// The stop is held until the stop transaction has settled (3A.2).
METHOD PRIVATE Stop_Is_Held_Until_The_Transaction_Settles
VAR_INST
	rig			: FB_IagRig;
	nStep		: INT;
	nCycles		: UINT;
	nEdges		: UINT;
	bSeen		: BOOL;
	sTest		: STRING(80);
END_VAR
TEST('Stop_Is_Held_Until_The_Transaction_Settles');
sTest := 'Stop_Is_Held_Until_The_Transaction_Settles: ';
IF nStep >= 90 THEN
	RETURN;
END_IF
rig.Scan();
nCycles := nCycles + 1;
CASE nStep OF
0:	// wait for the clock, then power on
	IF rig.ClockValid THEN
		rig.fbTel.Init();
		nStep := 10;
		nCycles := 0;
	ELSIF nCycles > 2000 THEN
		AssertTrue(Condition := FALSE, Message := 'the astronomical clock never became valid');
		F_Note(bFailed := TRUE, sText := CONCAT(sTest, 'the astronomical clock never became valid'));
		nStep := 99;
		TEST_FINISHED();
	END_IF
10:	// wait until the startup has finished (READY_STATE 1.0)
	IF rig.Online THEN
		rig.fbTel.Slew(fAzimuth := 180.0, fAltitude := 45.0);
		nStep := 20;
		nCycles := 0;
	ELSIF nCycles > 1500 THEN
		AssertTrue(Condition := FALSE, Message := 'the mock telescope did not reach READY_STATE 1.0');
		F_Note(bFailed := TRUE, sText := CONCAT(sTest, 'the mock telescope did not reach READY_STATE 1.0'));
		nStep := 99;
		TEST_FINISHED();
	END_IF
20:	// an axis is moving
	IF rig.fbHa.MoveAxis OR rig.fbDec.MoveAxis THEN
		nCycles := 0;
		nStep := 30;
	ELSIF nCycles > 300 THEN
		AssertTrue(Condition := FALSE, Message := 'the slew did not start an axis move');
		F_Note(bFailed := TRUE, sText := CONCAT(sTest, 'the slew did not start an axis move'));
		nStep := 99;
		TEST_FINISHED();
	END_IF
30:
	IF nCycles >= 5 THEN
		rig.fbTel.Stop();
		nStep := 40;
		nCycles := 0;
	END_IF
40:	// the stop is held while the axis is stopping, and released only when the transaction has settled
	IF nCycles = 2 THEN
		AssertTrue(Condition := rig.fbTel.bStopActive, Message := 'the stop is still held two scans after the command');
		F_Note(bFailed := NOT (rig.fbTel.bStopActive), sText := CONCAT(sTest, 'the stop is still held two scans after the command'));
	END_IF
	IF NOT rig.fbTel.bStopActive THEN
		AssertTrue(Condition := rig.fbTel.bSettled, Message := 'released only when settled');
		F_Note(bFailed := NOT (rig.fbTel.bSettled), sText := CONCAT(sTest, 'released only when settled'));
		nStep := 99;
		TEST_FINISHED();
	ELSIF nCycles > 400 THEN
		AssertTrue(Condition := FALSE, Message := 'the stop did not settle');
		F_Note(bFailed := TRUE, sText := CONCAT(sTest, 'the stop did not settle'));
		nStep := 99;
		TEST_FINISHED();
	END_IF
END_CASE
END_METHOD

// A goto and a home that are both pending when the stop comes are both cleared (3A.3).
METHOD PRIVATE Stop_Clears_Every_Pending_Move
VAR_INST
	rig			: FB_IagRig;
	nStep		: INT;
	nCycles		: UINT;
	nEdges		: UINT;
	bSeen		: BOOL;
	sTest		: STRING(80);
END_VAR
TEST('Stop_Clears_Every_Pending_Move');
sTest := 'Stop_Clears_Every_Pending_Move: ';
IF nStep >= 90 THEN
	RETURN;
END_IF
rig.Scan();
nCycles := nCycles + 1;
CASE nStep OF
0:	// wait for the clock, then power on
	IF rig.ClockValid THEN
		rig.fbTel.Init();
		nStep := 10;
		nCycles := 0;
	ELSIF nCycles > 2000 THEN
		AssertTrue(Condition := FALSE, Message := 'the astronomical clock never became valid');
		F_Note(bFailed := TRUE, sText := CONCAT(sTest, 'the astronomical clock never became valid'));
		nStep := 99;
		TEST_FINISHED();
	END_IF
10:	// wait until the startup has finished (READY_STATE 1.0)
	IF rig.Online THEN
		rig.fbTel.Track(fRightAscension := 100.0, fDeclination := 30.0);
		rig.fbTel.Home();
		rig.fbTel.Stop();
		nStep := 20;
		nCycles := 0;
	ELSIF nCycles > 1500 THEN
		AssertTrue(Condition := FALSE, Message := 'the mock telescope did not reach READY_STATE 1.0');
		F_Note(bFailed := TRUE, sText := CONCAT(sTest, 'the mock telescope did not reach READY_STATE 1.0'));
		nStep := 99;
		TEST_FINISHED();
	END_IF
20:	// one scan after the three commands
		AssertTrue(Condition := NOT rig.fbTel.bGotoActive, Message := 'the goto is gone');
		F_Note(bFailed := NOT (NOT rig.fbTel.bGotoActive), sText := CONCAT(sTest, 'the goto is gone'));
		AssertTrue(Condition := NOT rig.fbTel.bGoHomeActive, Message := 'the home is gone');
		F_Note(bFailed := NOT (NOT rig.fbTel.bGoHomeActive), sText := CONCAT(sTest, 'the home is gone'));
		nStep := 99;
		TEST_FINISHED();
END_CASE
END_METHOD

// A repeated stop does not send a second stop to an axis that is already stopping (3A.4).
METHOD PRIVATE Repeated_Stop_Restarts_Only_Moving_Axes
VAR_INST
	rig			: FB_IagRig;
	nStep		: INT;
	nCycles		: UINT;
	nEdges		: UINT;
	bSeen		: BOOL;
	sTest		: STRING(80);
END_VAR
TEST('Repeated_Stop_Restarts_Only_Moving_Axes');
sTest := 'Repeated_Stop_Restarts_Only_Moving_Axes: ';
IF nStep >= 90 THEN
	RETURN;
END_IF
rig.Scan();
nCycles := nCycles + 1;
CASE nStep OF
0:	// wait for the clock, then power on
	IF rig.ClockValid THEN
		rig.fbTel.Init();
		nStep := 10;
		nCycles := 0;
	ELSIF nCycles > 2000 THEN
		AssertTrue(Condition := FALSE, Message := 'the astronomical clock never became valid');
		F_Note(bFailed := TRUE, sText := CONCAT(sTest, 'the astronomical clock never became valid'));
		nStep := 99;
		TEST_FINISHED();
	END_IF
10:	// wait until the startup has finished (READY_STATE 1.0)
	IF rig.Online THEN
		rig.fbTel.Slew(fAzimuth := 180.0, fAltitude := 45.0);
		nStep := 20;
		nCycles := 0;
	ELSIF nCycles > 1500 THEN
		AssertTrue(Condition := FALSE, Message := 'the mock telescope did not reach READY_STATE 1.0');
		F_Note(bFailed := TRUE, sText := CONCAT(sTest, 'the mock telescope did not reach READY_STATE 1.0'));
		nStep := 99;
		TEST_FINISHED();
	END_IF
20:	// an axis is moving
	IF rig.fbHa.MoveAxis OR rig.fbDec.MoveAxis THEN
		nCycles := 0;
		nStep := 30;
	ELSIF nCycles > 300 THEN
		AssertTrue(Condition := FALSE, Message := 'the slew did not start an axis move');
		F_Note(bFailed := TRUE, sText := CONCAT(sTest, 'the slew did not start an axis move'));
		nStep := 99;
		TEST_FINISHED();
	END_IF
30:
	IF nCycles >= 5 THEN
		rig.fbTel.Stop();
		nStep := 35;
		nCycles := 0;
	END_IF
35:	// a second stop while the axis is already stopping (the stop reaches the axis in the third scan, the axis then reports Stopping)
	IF nCycles >= 3 THEN
		rig.fbTel.Stop();
		nStep := 40;
		nCycles := 0;
	END_IF
40:
	IF NOT rig.fbTel.bStopActive AND rig.fbTel.bStopped AND nCycles > 5 THEN
		AssertTrue(Condition := rig.fbHa.nStopEdges + rig.fbDec.nStopEdges = 1, Message := 'no second stop for an axis that was stopping');
		F_Note(bFailed := NOT (rig.fbHa.nStopEdges + rig.fbDec.nStopEdges = 1), sText := CONCAT(sTest, 'no second stop for an axis that was stopping'));
		nStep := 99;
		TEST_FINISHED();
	ELSIF nCycles > 400 THEN
		AssertTrue(Condition := FALSE, Message := 'the stop did not settle');
		F_Note(bFailed := TRUE, sText := CONCAT(sTest, 'the stop did not settle'));
		nStep := 99;
		TEST_FINISHED();
	END_IF
END_CASE
END_METHOD

// A park over a goto that is not dispatched yet runs a short abort stop, then the park (3A.5).
METHOD PRIVATE Park_Over_A_Waiting_Goto_Runs_A_Short_Abort_Stop
VAR_INST
	rig			: FB_IagRig;
	nStep		: INT;
	nCycles		: UINT;
	nEdges		: UINT;
	bSeen		: BOOL;
	sTest		: STRING(80);
END_VAR
TEST('Park_Over_A_Waiting_Goto_Runs_A_Short_Abort_Stop');
sTest := 'Park_Over_A_Waiting_Goto_Runs_A_Short_Abort_Stop: ';
IF nStep >= 90 THEN
	RETURN;
END_IF
rig.Scan();
nCycles := nCycles + 1;
CASE nStep OF
0:	// wait for the clock, then power on
	IF rig.ClockValid THEN
		rig.fbTel.Init();
		nStep := 10;
		nCycles := 0;
	ELSIF nCycles > 2000 THEN
		AssertTrue(Condition := FALSE, Message := 'the astronomical clock never became valid');
		F_Note(bFailed := TRUE, sText := CONCAT(sTest, 'the astronomical clock never became valid'));
		nStep := 99;
		TEST_FINISHED();
	END_IF
10:	// wait until the startup has finished (READY_STATE 1.0)
	IF rig.Online THEN
		rig.SetHorizon(-90.0);
		rig.SetSafeAltitude(-90.0);
		rig.fbTel.Track(fRightAscension := 100.0, fDeclination := 30.0);
		rig.fbTel.Park();
		nStep := 20;
		nCycles := 0;
	ELSIF nCycles > 1500 THEN
		AssertTrue(Condition := FALSE, Message := 'the mock telescope did not reach READY_STATE 1.0');
		F_Note(bFailed := TRUE, sText := CONCAT(sTest, 'the mock telescope did not reach READY_STATE 1.0'));
		nStep := 99;
		TEST_FINISHED();
	END_IF
20:	// the park preempted a goto that was not dispatched: the abort stop runs, then the park
	IF rig.fbTel.bMoveAbortPending THEN
		bSeen := TRUE;
	END_IF
	IF rig.fbTel.bIsParked THEN
		AssertTrue(Condition := bSeen, Message := 'the preemption ran the abort stop');
		F_Note(bFailed := NOT (bSeen), sText := CONCAT(sTest, 'the preemption ran the abort stop'));
		AssertTrue(Condition := NOT rig.fbTel.bGotoActive, Message := 'the goto is gone');
		F_Note(bFailed := NOT (NOT rig.fbTel.bGotoActive), sText := CONCAT(sTest, 'the goto is gone'));
		nStep := 99;
		TEST_FINISHED();
	ELSIF nCycles > 3000 THEN
		AssertTrue(Condition := FALSE, Message := 'the park did not finish');
		F_Note(bFailed := TRUE, sText := CONCAT(sTest, 'the park did not finish'));
		nStep := 99;
		TEST_FINISHED();
	END_IF
END_CASE
END_METHOD

END_FUNCTION_BLOCK

// ---- POUs/IagParkPowerReset_Tests.TcPOU
// Park, power-on and reset precedence of FB_TelescopeControl (IAG50cm), command model step 3B (BROTLib
// specs/plans/2026-11-09-iag50cm-command-model-unification.md). One rig per test, one Scan() per PLC cycle.
FUNCTION_BLOCK IagParkPowerReset_Tests EXTENDS TcUnit.FB_TestSuite
VAR
END_VAR

Park_During_Stop_Runs_After_Settle();
Stop_Drops_A_Park_Queued_Behind_A_Stop();
Init_During_Stop_Is_Refused();
Init_During_Park_Is_Refused();
Park_Right_After_Init_Aborts_The_PowerOn();
Init_Drops_A_Stale_Home();
Reset_At_Rest_Drops_A_Pending_Move();
Reset_During_Park_Keeps_The_Park();
Reset_Recovers_A_Stuck_Stop();

// A park sent during a stop runs when the stop has settled (D13).
METHOD PRIVATE Park_During_Stop_Runs_After_Settle
VAR_INST
	rig			: FB_IagRig;
	nStep		: INT;
	nCycles		: UINT;
	bSeen		: BOOL;
	sTest		: STRING(80);
END_VAR
TEST('Park_During_Stop_Runs_After_Settle');
sTest := 'Park_During_Stop_Runs_After_Settle: ';
IF nStep >= 90 THEN
	RETURN;
END_IF
rig.Scan();
nCycles := nCycles + 1;
CASE nStep OF
0:	// wait for the clock, then power on
	IF rig.ClockValid THEN
		rig.fbTel.Init();
		nStep := 10;
		nCycles := 0;
	ELSIF nCycles > 2000 THEN
		AssertTrue(Condition := FALSE, Message := 'the astronomical clock never became valid');
		F_Note(bFailed := TRUE, sText := CONCAT(sTest, 'the astronomical clock never became valid'));
		nStep := 99;
		TEST_FINISHED();
	END_IF
10:	// wait until the startup has finished (READY_STATE 1.0)
	IF rig.Online THEN
		rig.fbTel.Slew(fAzimuth := 180.0, fAltitude := 45.0);
		nStep := 20;
		nCycles := 0;
	ELSIF nCycles > 1500 THEN
		AssertTrue(Condition := FALSE, Message := 'the mock telescope did not reach READY_STATE 1.0');
		F_Note(bFailed := TRUE, sText := CONCAT(sTest, 'the mock telescope did not reach READY_STATE 1.0'));
		nStep := 99;
		TEST_FINISHED();
	END_IF
20:	// an axis is moving
	IF rig.fbHa.MoveAxis OR rig.fbDec.MoveAxis THEN
		nCycles := 0;
		nStep := 30;
	ELSIF nCycles > 300 THEN
		AssertTrue(Condition := FALSE, Message := 'the slew did not start an axis move');
		F_Note(bFailed := TRUE, sText := CONCAT(sTest, 'the slew did not start an axis move'));
		nStep := 99;
		TEST_FINISHED();
	END_IF
30:
	IF nCycles >= 5 THEN
		rig.fbTel.Stop();
		nStep := 35;
		nCycles := 0;
	END_IF
35:	// the stop runs: the park is queued behind it
	IF rig.fbTel.bStopActive THEN
		rig.fbTel.Park();
		nStep := 40;
		nCycles := 0;
	ELSIF nCycles > 10 THEN
		AssertTrue(Condition := FALSE, Message := 'the stop did not start');
		F_Note(bFailed := TRUE, sText := CONCAT(sTest, 'the stop did not start'));
		nStep := 99;
		TEST_FINISHED();
	END_IF
40:
		AssertTrue(Condition := rig.fbTel.bParkAfterStop, Message := 'the park is queued');
		F_Note(bFailed := NOT (rig.fbTel.bParkAfterStop), sText := CONCAT(sTest, 'the park is queued'));
		AssertTrue(Condition := NOT rig.fbTel.bParkActive, Message := 'the park does not run during the stop');
		F_Note(bFailed := NOT (NOT rig.fbTel.bParkActive), sText := CONCAT(sTest, 'the park does not run during the stop'));
	nStep := 50;
	nCycles := 0;
50:
	IF rig.fbTel.bIsParked THEN
		AssertTrue(Condition := NOT rig.fbTel.bParkAfterStop, Message := 'the queue is empty');
		F_Note(bFailed := NOT (NOT rig.fbTel.bParkAfterStop), sText := CONCAT(sTest, 'the queue is empty'));
		nStep := 99;
		TEST_FINISHED();
	ELSIF nCycles > 3000 THEN
		AssertTrue(Condition := FALSE, Message := 'the queued park did not run');
		F_Note(bFailed := TRUE, sText := CONCAT(sTest, 'the queued park did not run'));
		nStep := 99;
		TEST_FINISHED();
	END_IF
END_CASE
END_METHOD

// A stop clears a park that is queued behind a running stop (MONETcommon#213).
METHOD PRIVATE Stop_Drops_A_Park_Queued_Behind_A_Stop
VAR_INST
	rig			: FB_IagRig;
	nStep		: INT;
	nCycles		: UINT;
	bSeen		: BOOL;
	sTest		: STRING(80);
END_VAR
TEST('Stop_Drops_A_Park_Queued_Behind_A_Stop');
sTest := 'Stop_Drops_A_Park_Queued_Behind_A_Stop: ';
IF nStep >= 90 THEN
	RETURN;
END_IF
rig.Scan();
nCycles := nCycles + 1;
CASE nStep OF
0:	// wait for the clock, then power on
	IF rig.ClockValid THEN
		rig.fbTel.Init();
		nStep := 10;
		nCycles := 0;
	ELSIF nCycles > 2000 THEN
		AssertTrue(Condition := FALSE, Message := 'the astronomical clock never became valid');
		F_Note(bFailed := TRUE, sText := CONCAT(sTest, 'the astronomical clock never became valid'));
		nStep := 99;
		TEST_FINISHED();
	END_IF
10:	// wait until the startup has finished (READY_STATE 1.0)
	IF rig.Online THEN
		rig.fbTel.Slew(fAzimuth := 180.0, fAltitude := 45.0);
		nStep := 20;
		nCycles := 0;
	ELSIF nCycles > 1500 THEN
		AssertTrue(Condition := FALSE, Message := 'the mock telescope did not reach READY_STATE 1.0');
		F_Note(bFailed := TRUE, sText := CONCAT(sTest, 'the mock telescope did not reach READY_STATE 1.0'));
		nStep := 99;
		TEST_FINISHED();
	END_IF
20:	// an axis is moving
	IF rig.fbHa.MoveAxis OR rig.fbDec.MoveAxis THEN
		nCycles := 0;
		nStep := 30;
	ELSIF nCycles > 300 THEN
		AssertTrue(Condition := FALSE, Message := 'the slew did not start an axis move');
		F_Note(bFailed := TRUE, sText := CONCAT(sTest, 'the slew did not start an axis move'));
		nStep := 99;
		TEST_FINISHED();
	END_IF
30:
	IF nCycles >= 5 THEN
		rig.fbTel.Stop();
		nStep := 35;
		nCycles := 0;
	END_IF
35:
	IF rig.fbTel.bStopActive THEN
		rig.fbTel.Park();
		rig.fbTel.Stop();
		nStep := 40;
		nCycles := 0;
	ELSIF nCycles > 10 THEN
		AssertTrue(Condition := FALSE, Message := 'the stop did not start');
		F_Note(bFailed := TRUE, sText := CONCAT(sTest, 'the stop did not start'));
		nStep := 99;
		TEST_FINISHED();
	END_IF
40:
		AssertTrue(Condition := NOT rig.fbTel.bParkAfterStop, Message := 'the second stop dropped the queued park');
		F_Note(bFailed := NOT (NOT rig.fbTel.bParkAfterStop), sText := CONCAT(sTest, 'the second stop dropped the queued park'));
	nStep := 50;
	nCycles := 0;
50:	// the stop settles; no park follows
	IF nCycles >= 150 THEN
		AssertTrue(Condition := NOT rig.fbTel.bStopActive, Message := 'the stop is over');
		F_Note(bFailed := NOT (NOT rig.fbTel.bStopActive), sText := CONCAT(sTest, 'the stop is over'));
		AssertTrue(Condition := NOT rig.fbTel.bParkActive AND NOT rig.fbTel.bIsParked, Message := 'no park followed');
		F_Note(bFailed := NOT (NOT rig.fbTel.bParkActive AND NOT rig.fbTel.bIsParked), sText := CONCAT(sTest, 'no park followed'));
		nStep := 99;
		TEST_FINISHED();
	END_IF
END_CASE
END_METHOD

// A power-on during a stop is refused: a stop is not overridden by a power-on.
METHOD PRIVATE Init_During_Stop_Is_Refused
VAR_INST
	rig			: FB_IagRig;
	nStep		: INT;
	nCycles		: UINT;
	bSeen		: BOOL;
	sTest		: STRING(80);
END_VAR
TEST('Init_During_Stop_Is_Refused');
sTest := 'Init_During_Stop_Is_Refused: ';
IF nStep >= 90 THEN
	RETURN;
END_IF
rig.Scan();
nCycles := nCycles + 1;
CASE nStep OF
0:	// wait for the clock, then power on
	IF rig.ClockValid THEN
		rig.fbTel.Init();
		nStep := 10;
		nCycles := 0;
	ELSIF nCycles > 2000 THEN
		AssertTrue(Condition := FALSE, Message := 'the astronomical clock never became valid');
		F_Note(bFailed := TRUE, sText := CONCAT(sTest, 'the astronomical clock never became valid'));
		nStep := 99;
		TEST_FINISHED();
	END_IF
10:	// wait until the startup has finished (READY_STATE 1.0)
	IF rig.Online THEN
		rig.fbTel.Slew(fAzimuth := 180.0, fAltitude := 45.0);
		nStep := 20;
		nCycles := 0;
	ELSIF nCycles > 1500 THEN
		AssertTrue(Condition := FALSE, Message := 'the mock telescope did not reach READY_STATE 1.0');
		F_Note(bFailed := TRUE, sText := CONCAT(sTest, 'the mock telescope did not reach READY_STATE 1.0'));
		nStep := 99;
		TEST_FINISHED();
	END_IF
20:	// an axis is moving
	IF rig.fbHa.MoveAxis OR rig.fbDec.MoveAxis THEN
		nCycles := 0;
		nStep := 30;
	ELSIF nCycles > 300 THEN
		AssertTrue(Condition := FALSE, Message := 'the slew did not start an axis move');
		F_Note(bFailed := TRUE, sText := CONCAT(sTest, 'the slew did not start an axis move'));
		nStep := 99;
		TEST_FINISHED();
	END_IF
30:
	IF nCycles >= 5 THEN
		rig.fbTel.Stop();
		nStep := 35;
		nCycles := 0;
	END_IF
35:
	IF rig.fbTel.bStopActive THEN
		rig.fbTel.Init();
		nStep := 40;
		nCycles := 0;
	ELSIF nCycles > 10 THEN
		AssertTrue(Condition := FALSE, Message := 'the stop did not start');
		F_Note(bFailed := TRUE, sText := CONCAT(sTest, 'the stop did not start'));
		nStep := 99;
		TEST_FINISHED();
	END_IF
40:
		AssertTrue(Condition := rig.fbTel.nInitRefusedCount = 1, Message := 'the power-on was refused and counted');
		F_Note(bFailed := NOT (rig.fbTel.nInitRefusedCount = 1), sText := CONCAT(sTest, 'the power-on was refused and counted'));
		AssertTrue(Condition := NOT rig.fbTel.bPowerActive, Message := 'no power-on request');
		F_Note(bFailed := NOT (NOT rig.fbTel.bPowerActive), sText := CONCAT(sTest, 'no power-on request'));
		nStep := 99;
		TEST_FINISHED();
END_CASE
END_METHOD

// A power-on during a park is refused (the park is not cancelled by it any more).
METHOD PRIVATE Init_During_Park_Is_Refused
VAR_INST
	rig			: FB_IagRig;
	nStep		: INT;
	nCycles		: UINT;
	bSeen		: BOOL;
	sTest		: STRING(80);
END_VAR
TEST('Init_During_Park_Is_Refused');
sTest := 'Init_During_Park_Is_Refused: ';
IF nStep >= 90 THEN
	RETURN;
END_IF
rig.Scan();
nCycles := nCycles + 1;
CASE nStep OF
0:	// wait for the clock, then power on
	IF rig.ClockValid THEN
		rig.fbTel.Init();
		nStep := 10;
		nCycles := 0;
	ELSIF nCycles > 2000 THEN
		AssertTrue(Condition := FALSE, Message := 'the astronomical clock never became valid');
		F_Note(bFailed := TRUE, sText := CONCAT(sTest, 'the astronomical clock never became valid'));
		nStep := 99;
		TEST_FINISHED();
	END_IF
10:	// wait until the startup has finished (READY_STATE 1.0)
	IF rig.Online THEN
		rig.fbTel.Park();
		nStep := 20;
		nCycles := 0;
	ELSIF nCycles > 1500 THEN
		AssertTrue(Condition := FALSE, Message := 'the mock telescope did not reach READY_STATE 1.0');
		F_Note(bFailed := TRUE, sText := CONCAT(sTest, 'the mock telescope did not reach READY_STATE 1.0'));
		nStep := 99;
		TEST_FINISHED();
	END_IF
20:
	IF rig.fbTel.bParkActive THEN
		rig.fbTel.Init();
		nStep := 30;
		nCycles := 0;
	ELSIF nCycles > 10 THEN
		AssertTrue(Condition := FALSE, Message := 'the park did not start');
		F_Note(bFailed := TRUE, sText := CONCAT(sTest, 'the park did not start'));
		nStep := 99;
		TEST_FINISHED();
	END_IF
30:
		AssertTrue(Condition := rig.fbTel.nInitRefusedCount = 1, Message := 'the power-on was refused and counted');
		F_Note(bFailed := NOT (rig.fbTel.nInitRefusedCount = 1), sText := CONCAT(sTest, 'the power-on was refused and counted'));
		AssertTrue(Condition := NOT rig.fbTel.bPowerActive, Message := 'no power-on request');
		F_Note(bFailed := NOT (NOT rig.fbTel.bPowerActive), sText := CONCAT(sTest, 'no power-on request'));
		nStep := 99;
		TEST_FINISHED();
END_CASE
END_METHOD

// A park wins over a power-on that was requested in the same scan and not dispatched yet (D14).
METHOD PRIVATE Park_Right_After_Init_Aborts_The_PowerOn
VAR_INST
	rig			: FB_IagRig;
	nStep		: INT;
	nCycles		: UINT;
	bSeen		: BOOL;
	sTest		: STRING(80);
END_VAR
TEST('Park_Right_After_Init_Aborts_The_PowerOn');
sTest := 'Park_Right_After_Init_Aborts_The_PowerOn: ';
IF nStep >= 90 THEN
	RETURN;
END_IF
rig.Scan();
nCycles := nCycles + 1;
CASE nStep OF
0:	// Init() and Park() in one scan: the power-on is not dispatched yet, the park wins
	IF rig.ClockValid THEN
		rig.fbTel.Init();
		rig.fbTel.Park();
		nStep := 10;
		nCycles := 0;
	ELSIF nCycles > 2000 THEN
		AssertTrue(Condition := FALSE, Message := 'the astronomical clock never became valid');
		F_Note(bFailed := TRUE, sText := CONCAT(sTest, 'the astronomical clock never became valid'));
		nStep := 99;
		TEST_FINISHED();
	END_IF
10:
		AssertTrue(Condition := NOT rig.fbTel.bPowerActive, Message := 'the power-on was aborted by the park');
		F_Note(bFailed := NOT (NOT rig.fbTel.bPowerActive), sText := CONCAT(sTest, 'the power-on was aborted by the park'));
	nStep := 20;
	nCycles := 0;
20:
	IF rig.fbTel.bIsParked THEN
		AssertTrue(Condition := rig.fbTel.ReadyState <> 1.0, Message := 'the telescope did not come online');
		F_Note(bFailed := NOT (rig.fbTel.ReadyState <> 1.0), sText := CONCAT(sTest, 'the telescope did not come online'));
		nStep := 99;
		TEST_FINISHED();
	ELSIF nCycles > 3000 THEN
		AssertTrue(Condition := FALSE, Message := 'the park did not finish');
		F_Note(bFailed := TRUE, sText := CONCAT(sTest, 'the park did not finish'));
		nStep := 99;
		TEST_FINISHED();
	END_IF
END_CASE
END_METHOD

// A new power-on drops a stale home (the power-on homes itself at stage 100).
METHOD PRIVATE Init_Drops_A_Stale_Home
VAR_INST
	rig			: FB_IagRig;
	nStep		: INT;
	nCycles		: UINT;
	bSeen		: BOOL;
	sTest		: STRING(80);
END_VAR
TEST('Init_Drops_A_Stale_Home');
sTest := 'Init_Drops_A_Stale_Home: ';
IF nStep >= 90 THEN
	RETURN;
END_IF
rig.Scan();
nCycles := nCycles + 1;
CASE nStep OF
0:
	IF rig.ClockValid THEN
		rig.ForceGoHomeActive();	// a home left over from before
		rig.fbTel.Init();
		nStep := 10;
		nCycles := 0;
	ELSIF nCycles > 2000 THEN
		AssertTrue(Condition := FALSE, Message := 'the astronomical clock never became valid');
		F_Note(bFailed := TRUE, sText := CONCAT(sTest, 'the astronomical clock never became valid'));
		nStep := 99;
		TEST_FINISHED();
	END_IF
10:
		AssertTrue(Condition := rig.fbTel.bPowerActive, Message := 'the power-on runs');
		F_Note(bFailed := NOT (rig.fbTel.bPowerActive), sText := CONCAT(sTest, 'the power-on runs'));
		AssertTrue(Condition := NOT rig.fbTel.bGoHomeActive, Message := 'the stale home is gone');
		F_Note(bFailed := NOT (NOT rig.fbTel.bGoHomeActive), sText := CONCAT(sTest, 'the stale home is gone'));
		nStep := 99;
		TEST_FINISHED();
END_CASE
END_METHOD

// A reset without an error drops a pending move; the hardware part stays gated (Q1c).
METHOD PRIVATE Reset_At_Rest_Drops_A_Pending_Move
VAR_INST
	rig			: FB_IagRig;
	nStep		: INT;
	nCycles		: UINT;
	bSeen		: BOOL;
	sTest		: STRING(80);
END_VAR
TEST('Reset_At_Rest_Drops_A_Pending_Move');
sTest := 'Reset_At_Rest_Drops_A_Pending_Move: ';
IF nStep >= 90 THEN
	RETURN;
END_IF
rig.Scan();
nCycles := nCycles + 1;
CASE nStep OF
0:
	IF rig.ClockValid THEN
		rig.ForceSlewActive();	// a request that cannot run (the telescope is not on)
		rig.fbTel.Reset();
		nStep := 10;
		nCycles := 0;
	ELSIF nCycles > 2000 THEN
		AssertTrue(Condition := FALSE, Message := 'the astronomical clock never became valid');
		F_Note(bFailed := TRUE, sText := CONCAT(sTest, 'the astronomical clock never became valid'));
		nStep := 99;
		TEST_FINISHED();
	END_IF
10:
		AssertTrue(Condition := NOT rig.fbTel.bSlewActive, Message := 'the pending slew is dropped');
		F_Note(bFailed := NOT (NOT rig.fbTel.bSlewActive), sText := CONCAT(sTest, 'the pending slew is dropped'));
		AssertTrue(Condition := NOT rig.fbTel.bSafetyAckRequest, Message := 'no safety acknowledge without an error');
		F_Note(bFailed := NOT (NOT rig.fbTel.bSafetyAckRequest), sText := CONCAT(sTest, 'no safety acknowledge without an error'));
		AssertTrue(Condition := rig.fbHa.nResetEdges = 0 AND rig.fbDec.nResetEdges = 0, Message := 'no axis was reset');
		F_Note(bFailed := NOT (rig.fbHa.nResetEdges = 0 AND rig.fbDec.nResetEdges = 0), sText := CONCAT(sTest, 'no axis was reset'));
		nStep := 99;
		TEST_FINISHED();
END_CASE
END_METHOD

// A reset during a park does not stop it (its motion is wanted).
METHOD PRIVATE Reset_During_Park_Keeps_The_Park
VAR_INST
	rig			: FB_IagRig;
	nStep		: INT;
	nCycles		: UINT;
	bSeen		: BOOL;
	sTest		: STRING(80);
END_VAR
TEST('Reset_During_Park_Keeps_The_Park');
sTest := 'Reset_During_Park_Keeps_The_Park: ';
IF nStep >= 90 THEN
	RETURN;
END_IF
rig.Scan();
nCycles := nCycles + 1;
CASE nStep OF
0:	// wait for the clock, then power on
	IF rig.ClockValid THEN
		rig.fbTel.Init();
		nStep := 10;
		nCycles := 0;
	ELSIF nCycles > 2000 THEN
		AssertTrue(Condition := FALSE, Message := 'the astronomical clock never became valid');
		F_Note(bFailed := TRUE, sText := CONCAT(sTest, 'the astronomical clock never became valid'));
		nStep := 99;
		TEST_FINISHED();
	END_IF
10:	// wait until the startup has finished (READY_STATE 1.0)
	IF rig.Online THEN
		rig.fbTel.Park();
		nStep := 20;
		nCycles := 0;
	ELSIF nCycles > 1500 THEN
		AssertTrue(Condition := FALSE, Message := 'the mock telescope did not reach READY_STATE 1.0');
		F_Note(bFailed := TRUE, sText := CONCAT(sTest, 'the mock telescope did not reach READY_STATE 1.0'));
		nStep := 99;
		TEST_FINISHED();
	END_IF
20:
	IF rig.fbTel.bParkActive AND rig.fbTel.TCS_command = E_TCSCommand.park THEN
		rig.fbTel.Reset();
		nStep := 30;
		nCycles := 0;
	ELSIF nCycles > 300 THEN
		AssertTrue(Condition := FALSE, Message := 'the park did not start');
		F_Note(bFailed := TRUE, sText := CONCAT(sTest, 'the park did not start'));
		nStep := 99;
		TEST_FINISHED();
	END_IF
30:
	IF nCycles >= 3 THEN
		AssertTrue(Condition := rig.fbTel.bParkActive OR rig.fbTel.bIsParked, Message := 'the park goes on');
		F_Note(bFailed := NOT (rig.fbTel.bParkActive OR rig.fbTel.bIsParked), sText := CONCAT(sTest, 'the park goes on'));
		nStep := 40;
		nCycles := 0;
	END_IF
40:
	IF rig.fbTel.bIsParked THEN
		nStep := 99;
		TEST_FINISHED();
	ELSIF nCycles > 3000 THEN
		AssertTrue(Condition := FALSE, Message := 'the park did not finish');
		F_Note(bFailed := TRUE, sText := CONCAT(sTest, 'the park did not finish'));
		nStep := 99;
		TEST_FINISHED();
	END_IF
END_CASE
END_METHOD

// A reset recovers a stop that never gets its Done, without waiting for the 30 s timeout (D18).
METHOD PRIVATE Reset_Recovers_A_Stuck_Stop
VAR_INST
	rig			: FB_IagRig;
	nStep		: INT;
	nCycles		: UINT;
	bSeen		: BOOL;
	sTest		: STRING(80);
END_VAR
TEST('Reset_Recovers_A_Stuck_Stop');
sTest := 'Reset_Recovers_A_Stuck_Stop: ';
IF nStep >= 90 THEN
	RETURN;
END_IF
rig.Scan();
nCycles := nCycles + 1;
CASE nStep OF
0:	// wait for the clock, then power on
	IF rig.ClockValid THEN
		rig.fbTel.Init();
		nStep := 10;
		nCycles := 0;
	ELSIF nCycles > 2000 THEN
		AssertTrue(Condition := FALSE, Message := 'the astronomical clock never became valid');
		F_Note(bFailed := TRUE, sText := CONCAT(sTest, 'the astronomical clock never became valid'));
		nStep := 99;
		TEST_FINISHED();
	END_IF
10:	// wait until the startup has finished (READY_STATE 1.0)
	IF rig.Online THEN
		rig.SetStopWithoutDone(bHa := TRUE, bDec := TRUE);
		rig.fbTel.Slew(fAzimuth := 180.0, fAltitude := 45.0);
		nStep := 20;
		nCycles := 0;
	ELSIF nCycles > 1500 THEN
		AssertTrue(Condition := FALSE, Message := 'the mock telescope did not reach READY_STATE 1.0');
		F_Note(bFailed := TRUE, sText := CONCAT(sTest, 'the mock telescope did not reach READY_STATE 1.0'));
		nStep := 99;
		TEST_FINISHED();
	END_IF
20:	// an axis is moving
	IF rig.fbHa.MoveAxis OR rig.fbDec.MoveAxis THEN
		nCycles := 0;
		nStep := 30;
	ELSIF nCycles > 300 THEN
		AssertTrue(Condition := FALSE, Message := 'the slew did not start an axis move');
		F_Note(bFailed := TRUE, sText := CONCAT(sTest, 'the slew did not start an axis move'));
		nStep := 99;
		TEST_FINISHED();
	END_IF
30:
	IF nCycles >= 5 THEN
		rig.fbTel.Stop();
		nStep := 40;
		nCycles := 0;
	END_IF
40:	// the axes are at rest, the Done never comes: the stop is held
	IF rig.fbTel.bStopped AND nCycles > 6 THEN
		AssertTrue(Condition := rig.fbTel.bStopActive, Message := 'the stop is stuck');
		F_Note(bFailed := NOT (rig.fbTel.bStopActive), sText := CONCAT(sTest, 'the stop is stuck'));
		rig.fbTel.Reset();
		nStep := 50;
		nCycles := 0;
	ELSIF nCycles > 400 THEN
		AssertTrue(Condition := FALSE, Message := 'the axes did not come to rest');
		F_Note(bFailed := TRUE, sText := CONCAT(sTest, 'the axes did not come to rest'));
		nStep := 99;
		TEST_FINISHED();
	END_IF
50:	// the reset ends the stop at once, long before the 30 s timeout
	IF NOT rig.fbTel.bStopActive THEN
		AssertTrue(Condition := nCycles < 30, Message := 'released within a few scans');
		F_Note(bFailed := NOT (nCycles < 30), sText := CONCAT(sTest, 'released within a few scans'));
		AssertTrue(Condition := NOT rig.fbTel.bError, Message := 'no error');
		F_Note(bFailed := NOT (NOT rig.fbTel.bError), sText := CONCAT(sTest, 'no error'));
		nStep := 99;
		TEST_FINISHED();
	ELSIF nCycles > 100 THEN
		AssertTrue(Condition := FALSE, Message := 'the reset did not recover the stuck stop');
		F_Note(bFailed := TRUE, sText := CONCAT(sTest, 'the reset did not recover the stuck stop'));
		nStep := 99;
		TEST_FINISHED();
	END_IF
END_CASE
END_METHOD

END_FUNCTION_BLOCK

// ---- POUs/IagSupersede_Tests.TcPOU
// The latest move wins (supersede) in FB_TelescopeControl (IAG50cm), command model step 3C.1 (BROTLib
// specs/plans/2026-11-09-iag50cm-command-model-unification.md). The goto targets are not checked against the sky of the day
// (horizon and safe altitude -90). One rig per test, one Scan() per PLC cycle.
FUNCTION_BLOCK IagSupersede_Tests EXTENDS TcUnit.FB_TestSuite
VAR
END_VAR

Slew_During_Goto_Replaces_It();
Track_During_Goto_Retargets();
Home_During_Track_Stops_Then_Homes();

// A slew during a goto replaces it: the latest move wins (D6).
METHOD PRIVATE Slew_During_Goto_Replaces_It
VAR_INST
	rig			: FB_IagRig;
	nStep		: INT;
	nCycles		: UINT;
	bSeen		: BOOL;
	sTest		: STRING(80);
END_VAR
TEST('Slew_During_Goto_Replaces_It');
sTest := 'Slew_During_Goto_Replaces_It: ';
IF nStep >= 90 THEN
	RETURN;
END_IF
rig.Scan();
nCycles := nCycles + 1;
CASE nStep OF
0:	// wait for the clock, then power on
	IF rig.ClockValid THEN
		rig.fbTel.Init();
		nStep := 10;
		nCycles := 0;
	ELSIF nCycles > 2000 THEN
		AssertTrue(Condition := FALSE, Message := 'the astronomical clock never became valid');
		F_Note(bFailed := TRUE, sText := CONCAT(sTest, 'the astronomical clock never became valid'));
		nStep := 99;
		TEST_FINISHED();
	END_IF
10:	// wait until the startup has finished (READY_STATE 1.0)
	IF rig.Online THEN
		rig.SetHorizon(-90.0);
		rig.SetSafeAltitude(-90.0);
		rig.fbTel.Track(fRightAscension := 100.0, fDeclination := 30.0);
		nStep := 20;
		nCycles := 0;
	ELSIF nCycles > 1500 THEN
		AssertTrue(Condition := FALSE, Message := 'the mock telescope did not reach READY_STATE 1.0');
		F_Note(bFailed := TRUE, sText := CONCAT(sTest, 'the mock telescope did not reach READY_STATE 1.0'));
		nStep := 99;
		TEST_FINISHED();
	END_IF
20:	// the goto is moving an axis
	IF rig.fbHa.MoveAxis OR rig.fbDec.MoveAxis THEN
		nCycles := 0;
		nStep := 30;
	ELSIF nCycles > 300 THEN
		AssertTrue(Condition := FALSE, Message := 'the goto did not start an axis move');
		F_Note(bFailed := TRUE, sText := CONCAT(sTest, 'the goto did not start an axis move'));
		nStep := 99;
		TEST_FINISHED();
	END_IF
30:
	IF nCycles >= 5 THEN
		rig.fbTel.Slew(fAzimuth := 180.0, fAltitude := 45.0);
		nStep := 40;
		nCycles := 0;
	END_IF
40:	// the slew replaced the goto: the goto latch is gone, the abort stop runs, then the slew
	IF rig.fbTel.bMoveAbortPending THEN
		bSeen := TRUE;
	END_IF
	IF nCycles = 2 THEN
		AssertTrue(Condition := NOT rig.fbTel.bGotoActive, Message := 'the goto is gone');
		F_Note(bFailed := NOT (NOT rig.fbTel.bGotoActive), sText := CONCAT(sTest, 'the goto is gone'));
		AssertTrue(Condition := rig.fbTel.nCommandRejectCount = 0, Message := 'the slew was accepted');
		F_Note(bFailed := NOT (rig.fbTel.nCommandRejectCount = 0), sText := CONCAT(sTest, 'the slew was accepted'));
	END_IF
	IF nCycles > 5 AND NOT rig.fbTel.bSlewActive AND rig.fbTel.bStopped THEN
		AssertTrue(Condition := bSeen, Message := 'the replacement ran the abort stop');
		F_Note(bFailed := NOT (bSeen), sText := CONCAT(sTest, 'the replacement ran the abort stop'));
		AssertTrue(Condition := NOT rig.fbTel.bGotoActive, Message := 'the goto did not come back');
		F_Note(bFailed := NOT (NOT rig.fbTel.bGotoActive), sText := CONCAT(sTest, 'the goto did not come back'));
		nStep := 99;
		TEST_FINISHED();
	ELSIF nCycles > 3000 THEN
		AssertTrue(Condition := FALSE, Message := 'the slew did not finish');
		F_Note(bFailed := TRUE, sText := CONCAT(sTest, 'the slew did not finish'));
		nStep := 99;
		TEST_FINISHED();
	END_IF
END_CASE
END_METHOD

// A track during a goto retargets it through the abort stop (IAG#41).
METHOD PRIVATE Track_During_Goto_Retargets
VAR_INST
	rig			: FB_IagRig;
	nStep		: INT;
	nCycles		: UINT;
	bSeen		: BOOL;
	sTest		: STRING(80);
END_VAR
TEST('Track_During_Goto_Retargets');
sTest := 'Track_During_Goto_Retargets: ';
IF nStep >= 90 THEN
	RETURN;
END_IF
rig.Scan();
nCycles := nCycles + 1;
CASE nStep OF
0:	// wait for the clock, then power on
	IF rig.ClockValid THEN
		rig.fbTel.Init();
		nStep := 10;
		nCycles := 0;
	ELSIF nCycles > 2000 THEN
		AssertTrue(Condition := FALSE, Message := 'the astronomical clock never became valid');
		F_Note(bFailed := TRUE, sText := CONCAT(sTest, 'the astronomical clock never became valid'));
		nStep := 99;
		TEST_FINISHED();
	END_IF
10:	// wait until the startup has finished (READY_STATE 1.0)
	IF rig.Online THEN
		rig.SetHorizon(-90.0);
		rig.SetSafeAltitude(-90.0);
		rig.fbTel.Track(fRightAscension := 100.0, fDeclination := 30.0);
		nStep := 20;
		nCycles := 0;
	ELSIF nCycles > 1500 THEN
		AssertTrue(Condition := FALSE, Message := 'the mock telescope did not reach READY_STATE 1.0');
		F_Note(bFailed := TRUE, sText := CONCAT(sTest, 'the mock telescope did not reach READY_STATE 1.0'));
		nStep := 99;
		TEST_FINISHED();
	END_IF
20:	// the goto is moving an axis
	IF rig.fbHa.MoveAxis OR rig.fbDec.MoveAxis THEN
		nCycles := 0;
		nStep := 30;
	ELSIF nCycles > 300 THEN
		AssertTrue(Condition := FALSE, Message := 'the goto did not start an axis move');
		F_Note(bFailed := TRUE, sText := CONCAT(sTest, 'the goto did not start an axis move'));
		nStep := 99;
		TEST_FINISHED();
	END_IF
30:
	IF nCycles >= 5 THEN
		rig.fbTel.Track(fRightAscension := 110.0, fDeclination := 31.0);
		nStep := 40;
		nCycles := 0;
	END_IF
40:	// the second target replaces the first through the abort stop (IAG#41)
	IF rig.fbTel.bMoveAbortPending THEN
		bSeen := TRUE;
	END_IF
	IF nCycles > 5 AND rig.fbTel.TCS_command = E_TCSCommand.track THEN
		AssertTrue(Condition := bSeen, Message := 'the new target ran the abort stop');
		F_Note(bFailed := NOT (bSeen), sText := CONCAT(sTest, 'the new target ran the abort stop'));
		AssertTrue(Condition := ABS(rig.fbTel.fRightAscension - 110.0) < 0.001, Message := 'the new target is the one');
		F_Note(bFailed := NOT (ABS(rig.fbTel.fRightAscension - 110.0) < 0.001), sText := CONCAT(sTest, 'the new target is the one'));
		AssertTrue(Condition := rig.fbTel.nCommandRejectCount = 0, Message := 'nothing was rejected');
		F_Note(bFailed := NOT (rig.fbTel.nCommandRejectCount = 0), sText := CONCAT(sTest, 'nothing was rejected'));
		nStep := 99;
		TEST_FINISHED();
	ELSIF nCycles > 3000 THEN
		AssertTrue(Condition := FALSE, Message := 'the telescope did not reach the new target');
		F_Note(bFailed := TRUE, sText := CONCAT(sTest, 'the telescope did not reach the new target'));
		nStep := 99;
		TEST_FINISHED();
	END_IF
END_CASE
END_METHOD

// A home during tracking stops the tracking, then homes (IAG#72).
METHOD PRIVATE Home_During_Track_Stops_Then_Homes
VAR_INST
	rig			: FB_IagRig;
	nStep		: INT;
	nCycles		: UINT;
	bSeen		: BOOL;
	sTest		: STRING(80);
END_VAR
TEST('Home_During_Track_Stops_Then_Homes');
sTest := 'Home_During_Track_Stops_Then_Homes: ';
IF nStep >= 90 THEN
	RETURN;
END_IF
rig.Scan();
nCycles := nCycles + 1;
CASE nStep OF
0:	// wait for the clock, then power on
	IF rig.ClockValid THEN
		rig.fbTel.Init();
		nStep := 10;
		nCycles := 0;
	ELSIF nCycles > 2000 THEN
		AssertTrue(Condition := FALSE, Message := 'the astronomical clock never became valid');
		F_Note(bFailed := TRUE, sText := CONCAT(sTest, 'the astronomical clock never became valid'));
		nStep := 99;
		TEST_FINISHED();
	END_IF
10:	// wait until the startup has finished (READY_STATE 1.0)
	IF rig.Online THEN
		rig.SetHorizon(-90.0);
		rig.SetSafeAltitude(-90.0);
		rig.fbTel.Track(fRightAscension := 100.0, fDeclination := 30.0);
		nStep := 20;
		nCycles := 0;
	ELSIF nCycles > 1500 THEN
		AssertTrue(Condition := FALSE, Message := 'the mock telescope did not reach READY_STATE 1.0');
		F_Note(bFailed := TRUE, sText := CONCAT(sTest, 'the mock telescope did not reach READY_STATE 1.0'));
		nStep := 99;
		TEST_FINISHED();
	END_IF
20:	// wait until the mount tracks (the mock axes do not report isTracking: the track command is the sign)
	IF rig.fbTel.TCS_command = E_TCSCommand.track THEN
		rig.fbTel.Home();
		nStep := 30;
		nCycles := 0;
	ELSIF nCycles > 3000 THEN
		AssertTrue(Condition := FALSE, Message := 'the telescope did not track');
		F_Note(bFailed := TRUE, sText := CONCAT(sTest, 'the telescope did not track'));
		nStep := 99;
		TEST_FINISHED();
	END_IF
30:	// the home replaces the tracking: the abort stop ends the tracking, then the home runs (IAG#72)
	IF rig.fbTel.bMoveAbortPending THEN
		bSeen := TRUE;
	END_IF
	IF nCycles > 5 AND NOT rig.fbTel.bGoHomeActive AND rig.fbTel.bStopped THEN
		AssertTrue(Condition := bSeen, Message := 'the tracking was ended through the abort stop');
		F_Note(bFailed := NOT (bSeen), sText := CONCAT(sTest, 'the tracking was ended through the abort stop'));
		AssertTrue(Condition := rig.fbTel.TCS_command <> E_TCSCommand.track, Message := 'the telescope no longer tracks');
		F_Note(bFailed := NOT (rig.fbTel.TCS_command <> E_TCSCommand.track), sText := CONCAT(sTest, 'the telescope no longer tracks'));
		AssertTrue(Condition := rig.fbTel.nCommandRejectCount = 0, Message := 'the home was accepted');
		F_Note(bFailed := NOT (rig.fbTel.nCommandRejectCount = 0), sText := CONCAT(sTest, 'the home was accepted'));
		nStep := 99;
		TEST_FINISHED();
	ELSIF nCycles > 3000 THEN
		AssertTrue(Condition := FALSE, Message := 'the home did not finish');
		F_Note(bFailed := TRUE, sText := CONCAT(sTest, 'the home did not finish'));
		nStep := 99;
		TEST_FINISHED();
	END_IF
END_CASE
END_METHOD

END_FUNCTION_BLOCK

// ---- POUs/IagTelemetry_Tests.TcPOU
// Characterization of the telemetry of FB_TelescopeControl (IAG50cm#17, step 0 of specs/plans/2026-10-28-radec-telescope-control-migration-17.md):
// the field names and types that _SendTelemetryEquitorial (I:1868-2078) publishes, in order, and the values the clients
// depend on (pyBROT, BROTgui). The migration onto FB_RaDecTelescopeControl must not change them. FB_RecordingComm records
// the calls; the method is called once, directly, so the record holds exactly one telemetry run. The expected list was
// written from the code at IAG50cm develop 0df040e; where the code has an IF/ELSE with the same field in both branches the
// field is listed once.
FUNCTION_BLOCK IagTelemetry_Tests EXTENDS TcUnit.FB_TestSuite
VAR CONSTANT
	// kinds: 1 LREAL, 2 INT, 4 STRING (FB_RecordingComm)
	aExpectedNames : ARRAY[1..69] OF STRING(80) := [
		'TELESCOPE.READY_STATE',
		'TELESCOPE.MOTION_STATE',
		'TELESCOPE.INFO.NAME',
		'TELESCOPE.INFO.DIAMETER',
		'TELESCOPE.INFO.CABINET',
		'TELESCOPE.INFO.MANUFACTURER',
		'TELESCOPE.CONFIG.CAPABILITIES',
		'TELESCOPE.CONFIG.MOUNTOPTIONS',
		'TELESCOPE.CONFIG.MOUNT',
		'TELESCOPE.STATUS.GLOBAL',
		'TELESCOPE.STATUS.LOCAL_MODE',
		'OBJECT.INSTRUMENTAL.DEC',
		'OBJECT.INSTRUMENTAL.HA',
		'OBJECT.HORIZONTAL.ALT',
		'OBJECT.HORIZONTAL.AZ',
		'OBJECT.EQUATORIAL.EPOCH',
		'OBJECT.EQUATORIAL.EQUINOX',
		'OBJECT.EQUATORIAL.RA_PM',
		'OBJECT.EQUATORIAL.DEC_PM',
		'OBJECT.EQUATORIAL.RA_RATE',
		'OBJECT.EQUATORIAL.DEC_RATE',
		'OBJECT.EQUATORIAL.RA',
		'OBJECT.EQUATORIAL.DEC',
		'OBJECT.EQUATORIAL.HA_APPARENT',
		'OBJECT.EQUATORIAL.DEC_APPARENT',
		'POINTING.SLEWTIME',
		'POINTING.OFFSETS.HA',
		'POINTING.OFFSETS.DEC',
		'POSITION.LOCAL.SIDEREAL_TIME',
		'POSITION.LOCAL.JD',
		'POSITION.LOCAL.LATITUDE',
		'POSITION.LOCAL.LONGITUDE',
		'POSITION.LOCAL.HEIGHT',
		'POSITION.INSTRUMENTAL.DEC.POWER_STATE',
		'POSITION.INSTRUMENTAL.DEC.REFERENCED',
		'POSITION.INSTRUMENTAL.DEC.ERROR_STATE',
		'POSITION.INSTRUMENTAL.DEC.MOTION_STATE',
		'POSITION.INSTRUMENTAL.DEC.REALPOS',
		'POSITION.INSTRUMENTAL.DEC.CURRPOS',
		'POSITION.INSTRUMENTAL.DEC.TARGETPOS',
		'POSITION.INSTRUMENTAL.DEC.CURRSPEED',
		'POSITION.INSTRUMENTAL.DEC.TARGETDISTANCE',
		'POSITION.INSTRUMENTAL.DEC.OFFSET',
		'POSITION.INSTRUMENTAL.HA.POWER_STATE',
		'POSITION.INSTRUMENTAL.HA.REFERENCED',
		'POSITION.INSTRUMENTAL.HA.ERROR_STATE',
		'POSITION.INSTRUMENTAL.HA.MOTION_STATE',
		'POSITION.INSTRUMENTAL.HA.CURRPOS',
		'POSITION.INSTRUMENTAL.HA.REALPOS',
		'POSITION.INSTRUMENTAL.HA.TARGETPOS',
		'POSITION.INSTRUMENTAL.HA.CURRSPEED',
		'POSITION.INSTRUMENTAL.HA.TARGETDISTANCE',
		'POSITION.INSTRUMENTAL.HA.OFFSET',
		'POSITION.INSTRUMENTAL.FOCUS.POWER_STATE',
		'POSITION.INSTRUMENTAL.FOCUS.REFERENCED',
		'POSITION.INSTRUMENTAL.FOCUS.ERROR_STATE',
		'POSITION.INSTRUMENTAL.FOCUS.MOTION_STATE',
		'POSITION.INSTRUMENTAL.FOCUS.CURRPOS',
		'POSITION.INSTRUMENTAL.FOCUS.REALPOS',
		'POSITION.INSTRUMENTAL.FOCUS.TARGETPOS',
		'POSITION.INSTRUMENTAL.FOCUS.TARGETDISTANCE',
		'POSITION.INSTRUMENTAL.FOCUS.CURRSPEED',
		'POSITION.HORIZONTAL.ALT',
		'POSITION.HORIZONTAL.AZ',
		'POSITION.HORIZONTAL.DOME',
		'POSITION.EQUATORIAL.RA_ICRS',
		'POSITION.EQUATORIAL.DEC_ICRS',
		'POSITION.EQUATORIAL.HA_APPARENT',
		'POSITION.EQUATORIAL.DEC_APPARENT'];
	aExpectedKinds : ARRAY[1..69] OF INT := [1, 1, 4, 1, 4, 4, 2, 4, 4, 2, 2, 1, 1, 1, 1, 4, 4, 1, 1, 1, 1, 1, 1, 1, 1, 1, 1, 1, 1, 1, 1, 1, 1, 1, 1, 2, 2, 1, 1, 1, 1, 1, 1, 1, 1, 2, 2, 1, 1, 1, 1, 1, 1, 1, 1, 2, 2, 1, 1, 1, 1, 1, 1, 1, 1, 1, 1, 1, 1];
END_VAR

Telemetry_Field_Set_Is_Unchanged();
Telemetry_Offsets();
Telemetry_Estop_Global_1();
ReadyState_Is_Published_At_Power_On();

METHOD PRIVATE Telemetry_Field_Set_Is_Unchanged
VAR_INST
	rig			: FB_IagRig;
	nStep		: INT;
	nCycles		: UINT;
	sTest		: STRING(80);
	i			: INT;
	nFirstBad	: INT;
	nIdx		: INT;
END_VAR
TEST('Telemetry_Field_Set_Is_Unchanged');
sTest := 'Telemetry_Field_Set_Is_Unchanged: ';
IF nStep >= 90 THEN
	RETURN;
END_IF
rig.Scan();
nCycles := nCycles + 1;
CASE nStep OF
0:	// the telemetry method is called directly once the clock is valid, so nothing else publishes into the record
	IF rig.ClockValid THEN
		rig.fbComm.Start(sNameFilter := '');
		rig.fbTel._SendTelemetryEquitorial();
		rig.fbComm.Stop();
		nFirstBad := 0;
		FOR i := 1 TO 69 DO
			IF rig.fbComm.aNames[i] <> aExpectedNames[i] OR rig.fbComm.aKinds[i] <> aExpectedKinds[i] THEN
				nFirstBad := i;
				EXIT;
			END_IF
		END_FOR
		AssertEquals_INT(Expected := 69, Actual := rig.fbComm.nCount, Message := 'number of published fields');
		F_Note(bFailed := rig.fbComm.nCount <> 69, sText := CONCAT(sTest, CONCAT('number of published fields: ', INT_TO_STRING(rig.fbComm.nCount))));
		AssertEquals_INT(Expected := 0, Actual := nFirstBad, Message := 'first field that differs in name or type (index)');
		IF nFirstBad > 0 THEN
			F_Note(bFailed := TRUE, sText := CONCAT(CONCAT(CONCAT(sTest, CONCAT('field ', INT_TO_STRING(nFirstBad))), CONCAT(' is ', rig.fbComm.aNames[nFirstBad])), CONCAT(', expected ', aExpectedNames[nFirstBad])));
		END_IF
		nStep := 99;
		TEST_FINISHED();
	ELSIF nCycles > 2000 THEN
		AssertTrue(Condition := FALSE, Message := 'the astronomical clock never became valid');
		F_Note(bFailed := TRUE, sText := CONCAT(sTest, 'the astronomical clock never became valid'));
		nStep := 99;
		TEST_FINISHED();
	END_IF
END_CASE
END_METHOD

METHOD PRIVATE Telemetry_Offsets
VAR_INST
	rig			: FB_IagRig;
	nStep		: INT;
	nCycles		: UINT;
	sTest		: STRING(80);
	i			: INT;
	nFirstBad	: INT;
	nIdx		: INT;
END_VAR
TEST('Telemetry_Offsets');
sTest := 'Telemetry_Offsets: ';
IF nStep >= 90 THEN
	RETURN;
END_IF
rig.Scan();
nCycles := nCycles + 1;
CASE nStep OF
0:	// the telemetry method is called directly once the clock is valid, so nothing else publishes into the record
	IF rig.ClockValid THEN
		rig.SetOffsets(fHourAngle := 0.01, fDeclination := -0.02);
		rig.fbComm.Start(sNameFilter := '');
		rig.fbTel._SendTelemetryEquitorial();
		rig.fbComm.Stop();
		nIdx := rig.fbComm.FindName('POSITION.INSTRUMENTAL.HA.OFFSET');
		AssertTrue(Condition := nIdx > 0, Message := 'HA.OFFSET is published');
		F_Note(bFailed := nIdx <= 0, sText := CONCAT(sTest, 'HA.OFFSET is published'));
		IF nIdx > 0 THEN
			AssertFalse(Condition := F_NoteNear(sTest, 0.01, rig.fbComm.aValues[nIdx], 1.0E-12), Message := 'HA.OFFSET value');
		END_IF
		nIdx := rig.fbComm.FindName('POSITION.INSTRUMENTAL.DEC.OFFSET');
		AssertTrue(Condition := nIdx > 0, Message := 'DEC.OFFSET is published');
		F_Note(bFailed := nIdx <= 0, sText := CONCAT(sTest, 'DEC.OFFSET is published'));
		IF nIdx > 0 THEN
			AssertFalse(Condition := F_NoteNear(sTest, -0.02, rig.fbComm.aValues[nIdx], 1.0E-12), Message := 'DEC.OFFSET value');
		END_IF
		// BROTLib's FB_RaDecTelescopeControl publishes the hour-angle offset under RA.OFFSET (F3 of the plan); IAG must not
		nIdx := rig.fbComm.FindName('POSITION.INSTRUMENTAL.RA.OFFSET');
		AssertEquals_INT(Expected := 0, Actual := nIdx, Message := 'no RA.OFFSET field');
		F_Note(bFailed := nIdx <> 0, sText := CONCAT(sTest, 'no RA.OFFSET field'));
		nStep := 99;
		TEST_FINISHED();
	ELSIF nCycles > 2000 THEN
		AssertTrue(Condition := FALSE, Message := 'the astronomical clock never became valid');
		F_Note(bFailed := TRUE, sText := CONCAT(sTest, 'the astronomical clock never became valid'));
		nStep := 99;
		TEST_FINISHED();
	END_IF
END_CASE
END_METHOD

METHOD PRIVATE Telemetry_Estop_Global_1
VAR_INST
	rig			: FB_IagRig;
	nStep		: INT;
	nCycles		: UINT;
	sTest		: STRING(80);
	i			: INT;
	nFirstBad	: INT;
	nIdx		: INT;
END_VAR
TEST('Telemetry_Estop_Global_1');
sTest := 'Telemetry_Estop_Global_1: ';
IF nStep >= 90 THEN
	RETURN;
END_IF
rig.Scan();
nCycles := nCycles + 1;
CASE nStep OF
0:	// the telemetry method is called directly once the clock is valid, so nothing else publishes into the record
	IF rig.ClockValid THEN
		rig.SetEstop(bValue := TRUE);
		rig.fbComm.Start(sNameFilter := 'TELESCOPE.STATUS.GLOBAL');
		rig.fbTel._SendTelemetryEquitorial();
		rig.fbComm.Stop();
		AssertEquals_INT(Expected := 1, Actual := rig.fbComm.nCount, Message := 'one STATUS.GLOBAL record');
		F_Note(bFailed := rig.fbComm.nCount <> 1, sText := CONCAT(sTest, 'one STATUS.GLOBAL record'));
		IF rig.fbComm.nCount >= 1 THEN
			AssertFalse(Condition := F_NoteNear(sTest, 1.0, rig.fbComm.aValues[1], 1.0E-12), Message := 'E-stop is STATUS.GLOBAL 1 (#14)');
		END_IF
		nStep := 99;
		TEST_FINISHED();
	ELSIF nCycles > 2000 THEN
		AssertTrue(Condition := FALSE, Message := 'the astronomical clock never became valid');
		F_Note(bFailed := TRUE, sText := CONCAT(sTest, 'the astronomical clock never became valid'));
		nStep := 99;
		TEST_FINISHED();
	END_IF
END_CASE
END_METHOD

METHOD PRIVATE ReadyState_Is_Published_At_Power_On
VAR_INST
	rig			: FB_IagRig;
	nStep		: INT;
	nCycles		: UINT;
	sTest		: STRING(80);
	i			: INT;
	nFirstBad	: INT;
	nIdx		: INT;
END_VAR
TEST('ReadyState_Is_Published_At_Power_On');
sTest := 'ReadyState_Is_Published_At_Power_On: ';
IF nStep >= 90 THEN
	RETURN;
END_IF
rig.Scan();
nCycles := nCycles + 1;
CASE nStep OF
0:	// wait for the clock, then record only READY_STATE (the telemetry timer and PublishDue both publish it) and power on
	IF rig.ClockValid THEN
		rig.fbComm.Start(sNameFilter := 'TELESCOPE.READY_STATE');
		rig.fbTel.Init();
		nStep := 10;
		nCycles := 0;
	ELSIF nCycles > 2000 THEN
		AssertTrue(Condition := FALSE, Message := 'the astronomical clock never became valid');
		F_Note(bFailed := TRUE, sText := CONCAT(sTest, 'the astronomical clock never became valid'));
		nStep := 99;
		TEST_FINISHED();
	END_IF
10:	// READY_STATE 1.0 reached
	IF rig.Online THEN
		nStep := 20;
		nCycles := 0;
	ELSIF nCycles > 1500 THEN
		AssertTrue(Condition := FALSE, Message := 'the mock telescope did not reach READY_STATE 1.0');
		F_Note(bFailed := TRUE, sText := CONCAT(sTest, 'the mock telescope did not reach READY_STATE 1.0'));
		nStep := 99;
		TEST_FINISHED();
	END_IF
20:	// a few more scans so a publish on the change can come out (PublishDue, I:1023-1025)
	IF nCycles >= 10 THEN
		rig.fbComm.Stop();
		AssertTrue(Condition := rig.fbComm.nCount >= 1, Message := 'READY_STATE was published');
		F_Note(bFailed := rig.fbComm.nCount < 1, sText := CONCAT(sTest, 'READY_STATE was published'));
		IF rig.fbComm.nCount >= 1 THEN
			AssertEquals_INT(Expected := 1, Actual := rig.fbComm.aKinds[rig.fbComm.nCount], Message := 'published as LREAL');
			F_Note(bFailed := rig.fbComm.aKinds[rig.fbComm.nCount] <> 1, sText := CONCAT(sTest, 'published as LREAL'));
			AssertFalse(Condition := F_NoteNear(sTest, 1.0, rig.fbComm.aValues[rig.fbComm.nCount], 1.0E-12), Message := 'the last READY_STATE is 1.0');
		END_IF
		nStep := 99;
		TEST_FINISHED();
	END_IF
END_CASE
END_METHOD

END_FUNCTION_BLOCK

// ---- POUs/IagCoordinates_Tests.TcPOU
// Hand-value checks of FB_IagCoordinatesLegacy, the frozen coordinate chain of IAG50cm's FB_TelescopeControl (IAG50cm#17,
// step 0 of specs/plans/2026-10-28-radec-telescope-control-migration-17.md), so that the oracle is known to be sane before
// BROTLib's FB_RaDecCoordinates is compared against it (step 4). Site: the IAG 50 cm, JD 2461000.5. The expected values
// are geometry (zenith, meridian, pole), round trips between the two AstroBROT directions, and the sign and size of the
// offsets; tolerances are 0.01 deg where refraction or the frame could move the value, and written before the first CI run.
FUNCTION_BLOCK IagCoordinates_Tests EXTENDS TcUnit.FB_TestSuite
VAR
END_VAR

Current_At_The_Zenith_Is_90();
Current_On_The_Meridian_South();
Current_Near_The_Pole();
Current_Icrs_Roundtrips_Through_Target();
Corrected_Equals_Raw_Without_Offsets();
Offsets_Shift_The_Corrected_Position();
Inversion_Is_Held_When_Invalid();
Slew_Target_South_At_45();
Target_Below_The_Horizon();
Time_Offset_Shifts_The_Hour_Angle();

// HA 0 and Dec = latitude is the zenith. Raw current position (no refraction): elevation 90 within 0.01 deg.
METHOD PRIVATE Current_At_The_Zenith_Is_90
VAR
	fbA			: FB_IagCoordinatesLegacy;
	fbB			: FB_IagCoordinatesLegacy;
	sTest		: STRING(80);
	fDiff		: LREAL;
	bNote		: BOOL;
END_VAR
TEST('Current_At_The_Zenith_Is_90');
sTest := 'Current_At_The_Zenith_Is_90: ';
fbA.fJd := 2461000.5;
fbA.fLongitude := 9.9452433;
fbA.fLatitude := 51.5592378;
fbA.fAltitude := 100.0;
fbB.fJd := 2461000.5;
fbB.fLongitude := 9.9452433;
fbB.fLatitude := 51.5592378;
fbB.fAltitude := 100.0;
fbA.fHourAngleCurrent := 0.0;
fbA.fDeclinationCurrent := 51.5592378;
fbA();
AssertEquals_LREAL(Expected := 90.0, Actual := fbA.fElevationCurrent, Delta := 0.01, Message := 'elevation at the zenith');
bNote := F_NoteNear(CONCAT(sTest, 'elevation at the zenith'), 90.0, fbA.fElevationCurrent, 0.01);
TEST_FINISHED();
END_METHOD

// HA 0, Dec 0: culminates south at geometric elevation 90 - latitude = 38.44 deg, azimuth 180. The elevation of the current
// position (refract_to_observed := FALSE) is lower than the geometric one by the refraction (CI measured 38.4207, 0.020 deg
// less; Bennett's formula gives 0.021 deg at that height), so the tolerance is 0.05 deg.
METHOD PRIVATE Current_On_The_Meridian_South
VAR
	fbA			: FB_IagCoordinatesLegacy;
	fbB			: FB_IagCoordinatesLegacy;
	sTest		: STRING(80);
	fDiff		: LREAL;
	bNote		: BOOL;
END_VAR
TEST('Current_On_The_Meridian_South');
sTest := 'Current_On_The_Meridian_South: ';
fbA.fJd := 2461000.5;
fbA.fLongitude := 9.9452433;
fbA.fLatitude := 51.5592378;
fbA.fAltitude := 100.0;
fbB.fJd := 2461000.5;
fbB.fLongitude := 9.9452433;
fbB.fLatitude := 51.5592378;
fbB.fAltitude := 100.0;
fbA.fHourAngleCurrent := 0.0;
fbA.fDeclinationCurrent := 0.0;
fbA();
AssertEquals_LREAL(Expected := 90.0 - 51.5592378, Actual := fbA.fElevationCurrent, Delta := 0.05, Message := 'elevation');
bNote := F_NoteNear(CONCAT(sTest, 'elevation'), 90.0 - 51.5592378, fbA.fElevationCurrent, 0.05);
AssertEquals_LREAL(Expected := 180.0, Actual := fbA.fAzimuthCurrent, Delta := 0.05, Message := 'azimuth');
bNote := F_NoteNear(CONCAT(sTest, 'azimuth'), 180.0, fbA.fAzimuthCurrent, 0.05);
TEST_FINISHED();
END_METHOD

// HA 0, Dec 89.9: north of the zenith on the meridian, geometric elevation 90 - (89.9 - latitude) = 51.66 deg; CI measured
// 51.6464 (0.013 deg less, the refraction again, Bennett 0.013 deg), so the tolerance is 0.05 deg.
METHOD PRIVATE Current_Near_The_Pole
VAR
	fbA			: FB_IagCoordinatesLegacy;
	fbB			: FB_IagCoordinatesLegacy;
	sTest		: STRING(80);
	fDiff		: LREAL;
	bNote		: BOOL;
END_VAR
TEST('Current_Near_The_Pole');
sTest := 'Current_Near_The_Pole: ';
fbA.fJd := 2461000.5;
fbA.fLongitude := 9.9452433;
fbA.fLatitude := 51.5592378;
fbA.fAltitude := 100.0;
fbB.fJd := 2461000.5;
fbB.fLongitude := 9.9452433;
fbB.fLatitude := 51.5592378;
fbB.fAltitude := 100.0;
fbA.fHourAngleCurrent := 0.0;
fbA.fDeclinationCurrent := 89.9;
fbA();
AssertEquals_LREAL(Expected := 90.0 - (89.9 - 51.5592378), Actual := fbA.fElevationCurrent, Delta := 0.05, Message := 'elevation');
bNote := F_NoteNear(CONCAT(sTest, 'elevation'), 90.0 - (89.9 - 51.5592378), fbA.fElevationCurrent, 0.05);
TEST_FINISHED();
END_METHOD

// HA/Dec of the axes -> ICRS (current path) -> apparent HA/Dec of that target (target path): the inverse of each other.
METHOD PRIVATE Current_Icrs_Roundtrips_Through_Target
VAR
	fbA			: FB_IagCoordinatesLegacy;
	fbB			: FB_IagCoordinatesLegacy;
	sTest		: STRING(80);
	fDiff		: LREAL;
	bNote		: BOOL;
END_VAR
TEST('Current_Icrs_Roundtrips_Through_Target');
sTest := 'Current_Icrs_Roundtrips_Through_Target: ';
fbA.fJd := 2461000.5;
fbA.fLongitude := 9.9452433;
fbA.fLatitude := 51.5592378;
fbA.fAltitude := 100.0;
fbB.fJd := 2461000.5;
fbB.fLongitude := 9.9452433;
fbB.fLatitude := 51.5592378;
fbB.fAltitude := 100.0;
fbA.fHourAngleCurrent := 30.0;
fbA.fDeclinationCurrent := 40.0;
fbA();
fbB.fRightAscension := fbA.fRightAscensionCurrentICRS;
fbB.fDeclination := fbA.fDeclinationCurrentICRS;
fbB();
AssertEquals_LREAL(Expected := 30.0, Actual := fbB.fHourAngleApparent, Delta := 0.001, Message := 'hour angle');
bNote := F_NoteNear(CONCAT(sTest, 'hour angle'), 30.0, fbB.fHourAngleApparent, 0.001);
AssertEquals_LREAL(Expected := 40.0, Actual := fbB.fDeclinationApparent, Delta := 0.001, Message := 'declination');
bNote := F_NoteNear(CONCAT(sTest, 'declination'), 40.0, fbB.fDeclinationApparent, 0.001);
TEST_FINISHED();
END_METHOD

// No offset and a zero inversion: the corrected ICRS position is the raw one, exactly.
METHOD PRIVATE Corrected_Equals_Raw_Without_Offsets
VAR
	fbA			: FB_IagCoordinatesLegacy;
	fbB			: FB_IagCoordinatesLegacy;
	sTest		: STRING(80);
	fDiff		: LREAL;
	bNote		: BOOL;
END_VAR
TEST('Corrected_Equals_Raw_Without_Offsets');
sTest := 'Corrected_Equals_Raw_Without_Offsets: ';
fbA.fJd := 2461000.5;
fbA.fLongitude := 9.9452433;
fbA.fLatitude := 51.5592378;
fbA.fAltitude := 100.0;
fbB.fJd := 2461000.5;
fbB.fLongitude := 9.9452433;
fbB.fLatitude := 51.5592378;
fbB.fAltitude := 100.0;
fbA.fHourAngleCurrent := 30.0;
fbA.fDeclinationCurrent := 40.0;
fbA.bPointingInversionValid := TRUE;
fbA();
AssertEquals_LREAL(Expected := fbA.fRightAscensionCurrentICRS, Actual := fbA.fRightAscensionCurrentICRScorr, Delta := 1.0E-9, Message := 'RA');
bNote := F_NoteNear(CONCAT(sTest, 'RA'), fbA.fRightAscensionCurrentICRS, fbA.fRightAscensionCurrentICRScorr, 1.0E-9);
AssertEquals_LREAL(Expected := fbA.fDeclinationCurrentICRS, Actual := fbA.fDeclinationCurrentICRScorr, Delta := 1.0E-9, Message := 'Dec');
bNote := F_NoteNear(CONCAT(sTest, 'Dec'), fbA.fDeclinationCurrentICRS, fbA.fDeclinationCurrentICRScorr, 1.0E-9);
AssertEquals_LREAL(Expected := fbA.fElevationCurrent, Actual := fbA.fElevationCurrentSky, Delta := 1.0E-9, Message := 'sky elevation');
bNote := F_NoteNear(CONCAT(sTest, 'sky elevation'), fbA.fElevationCurrent, fbA.fElevationCurrentSky, 1.0E-9);
TEST_FINISHED();
END_METHOD

// A declination offset of 0.1 deg lowers the corrected Dec by 0.1 deg; an hour-angle offset of 0.05 deg on the sky moves the
// corrected RA by 0.05 / COS(Dec apparent) (F_HourAngleOffsetOnAxis), the sign being RA = LST - HA.
METHOD PRIVATE Offsets_Shift_The_Corrected_Position
VAR
	fbA			: FB_IagCoordinatesLegacy;
	fbB			: FB_IagCoordinatesLegacy;
	sTest		: STRING(80);
	fDiff		: LREAL;
	bNote		: BOOL;
	fRaShift	: LREAL;
END_VAR
TEST('Offsets_Shift_The_Corrected_Position');
sTest := 'Offsets_Shift_The_Corrected_Position: ';
fbA.fJd := 2461000.5;
fbA.fLongitude := 9.9452433;
fbA.fLatitude := 51.5592378;
fbA.fAltitude := 100.0;
fbB.fJd := 2461000.5;
fbB.fLongitude := 9.9452433;
fbB.fLatitude := 51.5592378;
fbB.fAltitude := 100.0;
fbA.fHourAngleCurrent := 30.0;
fbA.fDeclinationCurrent := 40.0;
fbA.fDeclinationOffset := 0.1;
fbA.fHourAngleOffset := 0.05;
fbA.fRightAscension := 100.0;
fbA.fDeclination := 40.0;
fbA();
AssertEquals_LREAL(Expected := -0.1, Actual := fbA.fDeclinationCurrentICRScorr - fbA.fDeclinationCurrentICRS, Delta := 0.001, Message := 'Dec shift');
bNote := F_NoteNear(CONCAT(sTest, 'Dec shift'), -0.1, fbA.fDeclinationCurrentICRScorr - fbA.fDeclinationCurrentICRS, 0.001);
fRaShift := fbA.fRightAscensionCurrentICRScorr - fbA.fRightAscensionCurrentICRS;
IF fRaShift > 180.0 THEN
	fRaShift := fRaShift - 360.0;
ELSIF fRaShift < -180.0 THEN
	fRaShift := fRaShift + 360.0;
END_IF
AssertEquals_LREAL(Expected := F_HourAngleOffsetOnAxis(0.05, fbA.fDeclinationApparent), Actual := fRaShift, Delta := 0.01, Message := 'RA shift');
bNote := F_NoteNear(CONCAT(sTest, 'RA shift'), F_HourAngleOffsetOnAxis(0.05, fbA.fDeclinationApparent), fRaShift, 0.01);
TEST_FINISHED();
END_METHOD

// FB_PointingModelInversion does not converge near the horizon (bValid FALSE): the last valid correction is kept (I:350-355)
// and used for the corrected position.
METHOD PRIVATE Inversion_Is_Held_When_Invalid
VAR
	fbA			: FB_IagCoordinatesLegacy;
	fbB			: FB_IagCoordinatesLegacy;
	sTest		: STRING(80);
	fDiff		: LREAL;
	bNote		: BOOL;
	fHaCorr	: LREAL;
END_VAR
TEST('Inversion_Is_Held_When_Invalid');
sTest := 'Inversion_Is_Held_When_Invalid: ';
fbA.fJd := 2461000.5;
fbA.fLongitude := 9.9452433;
fbA.fLatitude := 51.5592378;
fbA.fAltitude := 100.0;
fbB.fJd := 2461000.5;
fbB.fLongitude := 9.9452433;
fbB.fLatitude := 51.5592378;
fbB.fAltitude := 100.0;
fbA.fHourAngleCurrent := 30.0;
fbA.fDeclinationCurrent := 40.0;
fbA.fHourAngleInversionOffsetCalc := 0.5;
fbA.fDeclinationInversionOffsetCalc := 0.25;
fbA.bPointingInversionValid := TRUE;
fbA();
AssertEquals_LREAL(Expected := 0.5, Actual := fbA.fHourAngleInversionOffset, Delta := 1.0E-12, Message := 'held HA correction');
bNote := F_NoteNear(CONCAT(sTest, 'held HA correction'), 0.5, fbA.fHourAngleInversionOffset, 1.0E-12);
AssertEquals_LREAL(Expected := 0.25, Actual := fbA.fDeclinationInversionOffset, Delta := 1.0E-12, Message := 'held Dec correction');
bNote := F_NoteNear(CONCAT(sTest, 'held Dec correction'), 0.25, fbA.fDeclinationInversionOffset, 1.0E-12);
fHaCorr := fbA.fRightAscensionCurrentICRScorr;
fbA.fHourAngleInversionOffsetCalc := 9.0;
fbA.fDeclinationInversionOffsetCalc := 9.0;
fbA.bPointingInversionValid := FALSE;
fbA();
AssertEquals_LREAL(Expected := 0.5, Actual := fbA.fHourAngleInversionOffset, Delta := 1.0E-12, Message := 'HA correction kept');
bNote := F_NoteNear(CONCAT(sTest, 'HA correction kept'), 0.5, fbA.fHourAngleInversionOffset, 1.0E-12);
AssertEquals_LREAL(Expected := 0.25, Actual := fbA.fDeclinationInversionOffset, Delta := 1.0E-12, Message := 'Dec correction kept');
bNote := F_NoteNear(CONCAT(sTest, 'Dec correction kept'), 0.25, fbA.fDeclinationInversionOffset, 1.0E-12);
AssertEquals_LREAL(Expected := fHaCorr, Actual := fbA.fRightAscensionCurrentICRScorr, Delta := 1.0E-9, Message := 'corrected RA unchanged');
bNote := F_NoteNear(CONCAT(sTest, 'corrected RA unchanged'), fHaCorr, fbA.fRightAscensionCurrentICRScorr, 1.0E-9);
TEST_FINISHED();
END_METHOD

// Slew to azimuth 180, elevation 45 (alt_is_observed := FALSE, IAG50cm#3): on the meridian, Dec about latitude - 45 =
// 6.56 deg (J2000 and refraction move it by well under 0.5 deg), hour angle about 0.
METHOD PRIVATE Slew_Target_South_At_45
VAR
	fbA			: FB_IagCoordinatesLegacy;
	fbB			: FB_IagCoordinatesLegacy;
	sTest		: STRING(80);
	fDiff		: LREAL;
	bNote		: BOOL;
END_VAR
TEST('Slew_Target_South_At_45');
sTest := 'Slew_Target_South_At_45: ';
fbA.fJd := 2461000.5;
fbA.fLongitude := 9.9452433;
fbA.fLatitude := 51.5592378;
fbA.fAltitude := 100.0;
fbB.fJd := 2461000.5;
fbB.fLongitude := 9.9452433;
fbB.fLatitude := 51.5592378;
fbB.fAltitude := 100.0;
fbA.fElevation := 45.0;
fbA.fAzimuth := 180.0;
fbA();
AssertEquals_LREAL(Expected := 51.5592378 - 45.0, Actual := fbA.fDeclinationCalc, Delta := 0.5, Message := 'Dec');
bNote := F_NoteNear(CONCAT(sTest, 'Dec'), 51.5592378 - 45.0, fbA.fDeclinationCalc, 0.5);
AssertTrue(Condition := COS(fbA.fHourAngleCalc * 0.017453292519943295) > 0.9999, Message := 'hour angle about 0');
F_Note(bFailed := NOT (COS(fbA.fHourAngleCalc * 0.017453292519943295) > 0.9999), sText := CONCAT(sTest, CONCAT('hour angle about 0, got ', LREAL_TO_STRING(fbA.fHourAngleCalc))));
TEST_FINISHED();
END_METHOD

// Dec -60 never rises at 51.6 deg north (maximum elevation 90 - 51.56 - 60 = -21.6 deg): the target elevation is negative.
METHOD PRIVATE Target_Below_The_Horizon
VAR
	fbA			: FB_IagCoordinatesLegacy;
	fbB			: FB_IagCoordinatesLegacy;
	sTest		: STRING(80);
	fDiff		: LREAL;
	bNote		: BOOL;
END_VAR
TEST('Target_Below_The_Horizon');
sTest := 'Target_Below_The_Horizon: ';
fbA.fJd := 2461000.5;
fbA.fLongitude := 9.9452433;
fbA.fLatitude := 51.5592378;
fbA.fAltitude := 100.0;
fbB.fJd := 2461000.5;
fbB.fLongitude := 9.9452433;
fbB.fLatitude := 51.5592378;
fbB.fAltitude := 100.0;
fbA.fRightAscension := 100.0;
fbA.fDeclination := -60.0;
fbA();
AssertTrue(Condition := fbA.fElevationCalc < 0.0, Message := 'target below the horizon');
F_Note(bFailed := NOT (fbA.fElevationCalc < 0.0), sText := CONCAT(sTest, CONCAT('elevation ', LREAL_TO_STRING(fbA.fElevationCalc))));
TEST_FINISHED();
END_METHOD

// fTimeOffset is days added to the Julian date: half a day moves the hour angle by half a sidereal rotation, 180.49 deg.
METHOD PRIVATE Time_Offset_Shifts_The_Hour_Angle
VAR
	fbA			: FB_IagCoordinatesLegacy;
	fbB			: FB_IagCoordinatesLegacy;
	sTest		: STRING(80);
	fDiff		: LREAL;
	bNote		: BOOL;
END_VAR
TEST('Time_Offset_Shifts_The_Hour_Angle');
sTest := 'Time_Offset_Shifts_The_Hour_Angle: ';
fbA.fJd := 2461000.5;
fbA.fLongitude := 9.9452433;
fbA.fLatitude := 51.5592378;
fbA.fAltitude := 100.0;
fbB.fJd := 2461000.5;
fbB.fLongitude := 9.9452433;
fbB.fLatitude := 51.5592378;
fbB.fAltitude := 100.0;
fbA.fRightAscension := 100.0;
fbA.fDeclination := 20.0;
fbA();
fbB.fRightAscension := 100.0;
fbB.fDeclination := 20.0;
fbB.fTimeOffset := 0.5;
fbB();
fDiff := fbB.fHourAngleApparent - fbA.fHourAngleApparent;
WHILE fDiff < 0.0 DO
	fDiff := fDiff + 360.0;
END_WHILE
WHILE fDiff >= 360.0 DO
	fDiff := fDiff - 360.0;
END_WHILE
AssertEquals_LREAL(Expected := 180.4928, Actual := fDiff, Delta := 0.02, Message := 'hour angle shift');
bNote := F_NoteNear(CONCAT(sTest, 'hour angle shift'), 180.4928, fDiff, 0.02);
TEST_FINISHED();
END_METHOD

END_FUNCTION_BLOCK

// ---- POUs/FB_IagCoordinatesLegacy.TcPOU
// The coordinate chain of IAG50cm's FB_TelescopeControl as it is at IAG50cm develop 0df040e (FB_TelescopeControl.TcPOU
// lines 297-397 and 217-222 minus the clock), frozen into a block of its own: the oracle for IAG50cm#17 (step 0 of
// specs/plans/2026-10-28-radec-telescope-control-migration-17.md). The same AstroBROT calls in the same order with the
// same instances (the one fbEq2Hor is called three times, as in the telescope). Do not "improve" it: step 4 of the plan
// compares BROTLib's FB_RaDecCoordinates against this block. The pointing models stay in the telescope, so their
// results come in as inputs (fHourAngleInversionOffsetCalc/fDeclinationInversionOffsetCalc/bPointingInversionValid).
FUNCTION_BLOCK FB_IagCoordinatesLegacy
VAR_INPUT
	fJd								: LREAL;	// Julian date of the clock; the block adds fTimeOffset like the telescope
	fTimeOffset						: LREAL;
	fLongitude						: LREAL;	// telescopeConfig.longitude
	fLatitude						: LREAL;
	fAltitude						: LREAL;
	fRightAscension					: LREAL;	// target, ICRS degrees (TCS input)
	fDeclination					: LREAL;
	fElevation						: LREAL;	// slew target (TCS input)
	fAzimuth						: LREAL;
	fHourAngleCurrent				: LREAL;	// axis positions
	fDeclinationCurrent				: LREAL;
	fHourAngleOffset				: LREAL;	// user offsets
	fDeclinationOffset				: LREAL;
	fHourAngleInversionOffsetCalc	: LREAL;	// raw outputs of FB_PointingModelInversion this scan
	fDeclinationInversionOffsetCalc	: LREAL;
	bPointingInversionValid			: BOOL;
END_VAR
VAR_OUTPUT
	fHourAngleApparent				: LREAL;
	fDeclinationApparent			: LREAL;
	fElevationCalc					: LREAL;
	fAzimuthCalc					: LREAL;
	fRightAscensionCalc				: LREAL;
	fDeclinationCalc				: LREAL;
	fHourAngleCalc					: LREAL;
	fHourAngleInversionOffset		: LREAL;	// the last valid inversion correction
	fDeclinationInversionOffset		: LREAL;
	fRightAscensionCurrentICRS		: LREAL;
	fDeclinationCurrentICRS			: LREAL;
	fRightAscensionCurrentICRScorr	: LREAL;
	fDeclinationCurrentICRScorr		: LREAL;
	fElevationCurrent				: LREAL;
	fAzimuthCurrent					: LREAL;
	fElevationCurrentSky			: LREAL;
	fAzimuthCurrentSky				: LREAL;
END_VAR
VAR
	fbEq2Hor			: FB_EQ2HOR;
	fbHor2Eq			: FB_HOR2EQ;
	fbHaDec2RaDec		: FB_HADEC2RADEC;
	fbRaDec2HaDec		: FB_RADEC2HADEC;
END_VAR

// calculate fHourAngleApparent, fDeclinationApparent

fbRaDec2HaDec(
	ra := fRightAscension,
	dec := fDeclination,
	lon := fLongitude,
	JD := fJd + fTimeOffset,
	ha_out => fHourAngleApparent,
	dec_out => fDeclinationApparent);
// (and also horizontal coord. -> used for checking if target is on sky or in ground)
fbEq2Hor(
	ra := fRightAscension,
	dec := fDeclination,
	lon := fLongitude,
	lat := fLatitude,
	altitude := fAltitude,
	JD := fJd + fTimeOffset,
	refract_to_observed := TRUE,
	alt => fElevationCalc,
	az => fAzimuthCalc);

// calculate equatorial coordinates (used by Slew command, takes Alt/Az -> moves telescope)
fbHor2Eq(alt := fElevation,
		az := fAzimuth,
		jd := fJd+fTimeOffset,
		lat := fLatitude,
		lon := fLongitude,
		altitude := fAltitude,
		alt_is_observed := FALSE,
		ra => fRightAscensionCalc,
		dec => fDeclinationCalc,
		ha => fHourAngleCalc);
// (the pointing forward model sits here in the telescope; it does not feed back into these outputs)
// near the horizon the inversion is chaotic and does not converge (see FB_PointingModelInversion);
// keep reporting the last trustworthy correction rather than whatever garbage it would return
IF bPointingInversionValid THEN
	fHourAngleInversionOffset := fHourAngleInversionOffsetCalc;
	fDeclinationInversionOffset := fDeclinationInversionOffsetCalc;
END_IF
(*--------------------------------------------------------------*)
// transform from apparent to icrs

//current
fbHaDec2RaDec(
	ha := fHourAngleCurrent,
	dec := fDeclinationCurrent,
	jd := fJd+fTimeOffset,
	lon := fLongitude,
	ra_out => fRightAscensionCurrentICRS,
	dec_out => fDeclinationCurrentICRS);
//current corrected
fbHaDec2RaDec(
	ha := fHourAngleCurrent - fHourAngleInversionOffset - F_HourAngleOffsetOnAxis(fHourAngleOffset, fDeclinationApparent),
	dec := fDeclinationCurrent - fDeclinationInversionOffset- fDeclinationOffset,
	jd := fJd+fTimeOffset,
	lon := fLongitude,
	ra_out => fRightAscensionCurrentICRScorr,
	dec_out => fDeclinationCurrentICRScorr);
(*--------------------------------------------------------------*)
// to ALT AZ
fbEq2Hor(
	ra := fRightAscensionCurrentICRS,
	dec := fDeclinationCurrentICRS,
	lon := fLongitude,
	lat := fLatitude,
	altitude := fAltitude,
	refract_to_observed := FALSE,
	JD := fJd + fTimeOffset,
	alt => fElevationCurrent,
	az => fAzimuthCurrent);

fbEq2Hor(
	ra := fRightAscensionCurrentICRScorr,
	dec := fDeclinationCurrentICRScorr,
	lon := fLongitude,
	lat := fLatitude,
	altitude := fAltitude,
	refract_to_observed := FALSE,
	JD := fJd + fTimeOffset,
	alt => fElevationCurrentSky,
	az => fAzimuthCurrentSky);

END_FUNCTION_BLOCK
